{region 'Documentation'}
(*!
<summary>Checks inequality with the forbidden DT value.</summary>
*)
{endregion}
FUNCTION_BLOCK AssertNotEqual_DT EXTENDS AssertionBase
VAR_INPUT
    IN : DT; //! Actual value checked or observed by this Assertion.
    Expected : DT; //! Value that must differ from IN under this Assertion's comparison rules.
END_VAR

SUPER^();

{region 'Documentation'}
(*!
<summary>Evaluate the typed temporal relation and report higher-priority errors first.</summary>
*)
{endregion}
METHOD PROTECTED Assert
VAR
    Message : STRING(GVL_Constants.MessageLength);
    ExpectedText : STRING(GVL_Constants.AssertionValueLength);
    ActualText : STRING(GVL_Constants.AssertionValueLength);
END_VAR
IF NOT EvaluationActive THEN
    RETURN;
END_IF;

IF Result = E_Result.Error THEN
    RETURN;
END_IF;

IF Result = E_Result.Failed THEN
    RETURN;
END_IF;

IF IN = Expected THEN
    ExpectedText := DT_TO_STRING(Expected);
    ActualText := DT_TO_STRING(IN);
    Message := CONCAT('Assertion failed: values are equal but should differ. NotExpected = ',
        ExpectedText);
    Message := CONCAT(Message, ', Actual = ');
    Message := CONCAT(Message, ActualText);
    Message := CONCAT(Message, '.');
    Fail(Message := Message);
    RETURN;
END_IF;

Pass();
END_METHOD

END_FUNCTION_BLOCK

(* stored: Version 1.1.0.1
   POU AssertNotEqual_DT: Id {0d38f415-7a00-45c1-8d1a-c30f56200caa}, SpecialFunc None
   Folder Internal: Id {4bdaad28-45a5-4354-883f-bf8bc12bb92e}
   Method Assert: Id {9699f90d-5288-4661-b01b-2c1ac6b3ec50} *)
